(* IEC 61131-3 sources: SRCI_CLIENT_PLC/RobotLibrary/Library/Structures/Telegram/RobToPlc/Command, 2 files *)

(* ---- TelegramRobToPlcCommand.st ---- *)
{attribute 'pack_mode' := '1'}
// -------------------------------------------------------------------------
//  SRCI Robot Library
// -------------------------------------------------------------------------
//
//  Object:      TelegramPlcToRobMessage
//  Author:      Thorsten Brach
//  Date:        2024-11-02
//
//  Description:
//
//
//  Copyright:
//    (C) 2024 Thorsten Brach. All rights reserved
//             Licensed under the MIT License.
//
//  Disclaimer:
//    This project is provided without any guarantee and can be used for
//    private and commercial purposes. Any use is at the user’s
//    own risk and responsibility.
//
// -------------------------------------------------------------------------
TYPE TelegramRobToPlcCommand :
STRUCT
  /// Header
  Header  : TelegramRobToPlcCommandHeader;
  /// Payload
  Payload : ARRAY[0..RobotLibraryParameter.RESPONSE_PAYLOAD_MAX] OF BYTE;
END_STRUCT
END_TYPE

(* ---- TelegramRobToPlcCommandHeader.st ---- *)
{attribute 'pack_mode' := '1'}
// -------------------------------------------------------------------------
//  SRCI Robot Library
// -------------------------------------------------------------------------
//
//  Object:      TelegramPlcToRobMessageHeader
//  Author:      Thorsten Brach
//  Date:        2024-11-02
//
//  Description:
//
//
//  Copyright:
//    (C) 2024 Thorsten Brach. All rights reserved
//             Licensed under the MIT License.
//
//  Disclaimer:
//    This project is provided without any guarantee and can be used for
//    private and commercial purposes. Any use is at the user’s
//    own risk and responsibility.
//
// -------------------------------------------------------------------------
TYPE TelegramRobToPlcCommandHeader :
STRUCT
  /// Parameter squence
  ParSeq               : BYTE;
  /// message Staet
  State                : CmdMessageState;
  /// Alarm Message Severity
  AlarmMessageSeverity : SINT;
  /// Alarm Message Code
  AlarmMessageCode     : UINT;
END_STRUCT
END_TYPE
